// TIA Portal V21 export
// export: Created 2026-10-23T20:42:46.0665102Z, ExportSetting WithDefaults, DisplayName Totally Integrated Automation Portal, DisplayVersion V21 Update 1, DisplayName SINAMICS Startdrive Advanced, DisplayVersion V21 HF2, DisplayName SINAMICS Startdrive G110M, G120, G120C, G120D, G120P, G115D, DisplayVersion V21 HF2, DisplayName SINAMICS Startdrive G130, G150, S120, S150, G200, G220, S200, S210, S220, Innomotics MVD, DisplayVersion V21 HF2, DisplayName STEP 7 Professional, DisplayVersion V21 Update 1, DisplayName STEP 7 Safety, DisplayVersion V21, DisplayName Tech WebApplication, DisplayVersion V21, DisplayName WinCC Basic/Comfort/Advanced, DisplayVersion V21 Update 1, DisplayName WinCC Unified, DisplayVersion V21 Update 1
FUNCTION "FC_FbdLogic" : Void   // FC8, FBD
TITLE = FUP-Logik / FBD logic
{ S7_Optimized_Access := 'TRUE' }
VERSION : 0.1
// UND, ODER, XOR, Negation, Zuweisung, SR, RS und Flankenerkennung in FUP / AND, OR, XOR, negation, assignment, SR, RS and edge detection in FBD
// stored: AutoNumber true, IsIECCheckEnabled false, SetENOAutomatically false, UDAEnableTagReadback false
   VAR_INPUT
      InA : Bool;
      InB : Bool;
   END_VAR
   VAR_OUTPUT
      AndOut : Bool;
      OrOut : Bool;
      XorOut : Bool;
      NotOut : Bool;
      SrOut : Bool;
      RsOut : Bool;
      EdgeOut : Bool;
   END_VAR
   VAR_IN_OUT
      SrBit : Bool;
      RsBit : Bool;
      EdgeBit : Bool;
   END_VAR
   VAR_TEMP   // added for the SCL form of the ladder/FBD networks
      _w1 : Bool;
   END_VAR
BEGIN

REGION Network 1: UND / AND
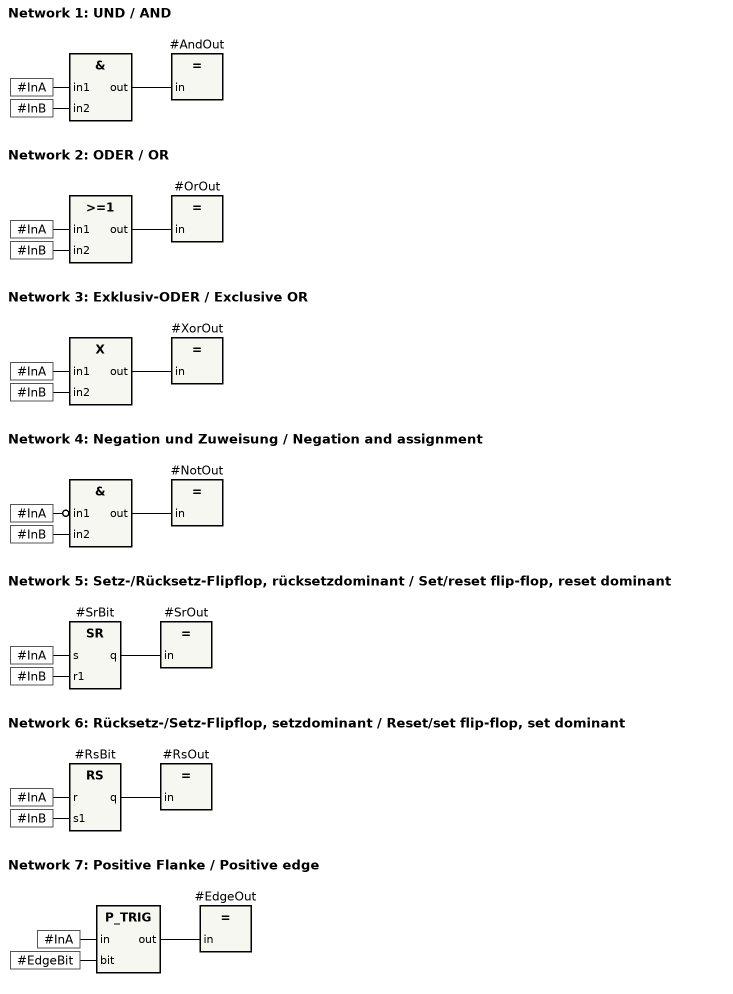
   #AndOut := #InA AND #InB;
END_REGION

REGION Network 2: ODER / OR
   #OrOut := #InA OR #InB;
END_REGION

REGION Network 3: Exklusiv-ODER / Exclusive OR
   #XorOut := #InA XOR #InB;
END_REGION

REGION Network 4: Negation und Zuweisung / Negation and assignment
   #NotOut := NOT #InA AND #InB;
END_REGION

REGION Network 5: Setz-/Rücksetz-Flipflop, rücksetzdominant / Set/reset flip-flop, reset dominant
   IF #InA THEN
       #SrBit := TRUE;   // SR flip-flop
   END_IF;
   IF #InB THEN #SrBit := FALSE; END_IF;
   #SrOut := #SrBit;
END_REGION

REGION Network 6: Rücksetz-/Setz-Flipflop, setzdominant / Reset/set flip-flop, set dominant
   IF #InA THEN
       #RsBit := FALSE;   // RS flip-flop
   END_IF;
   IF #InB THEN #RsBit := TRUE; END_IF;
   #RsOut := #RsBit;
END_REGION

REGION Network 7: Positive Flanke / Positive edge
   #_w1 := #InA AND NOT #EdgeBit;   // rising edge
   #EdgeBit := #InA;
   #EdgeOut := #_w1;
END_REGION
END_FUNCTION
